Fanuc KAREL source: KT00719.KL

PROGRAM KT00719
%NOLOCKGROUP
VAR
  P1: POSITION
  P2: POSITION
  OUT: INTEGER
BEGIN
  OUT = ARRAY_LEN(P1)
END KT00719
